TYPE ST_HomingResult :
STRUCT
	HomePos_Beta  : LREAL;   (* joint angle/position after homing *)
    HomePos_Theta  : LREAL;
    HomePos_R  : LREAL;
END_STRUCT
END_TYPE

(* stored: Version 1.1.0.1, ProductVersion 3.1.4024.15
   DUT ST_HomingResult: Id {37118aec-59c1-4ce7-8906-671357d16b92} *)
